(* IEC 61131-3 sources: SRCI_CLIENT_PLC/RobotLibrary/Library/Structures/DatenAndTime, 4 files *)

(* ---- IEC_DATE.st ---- *)
/// Date in the format days since 1990.01.01
TYPE IEC_DATE : UINT;
// -------------------------------------------------------------------------
//  SRCI Robot Library
// -------------------------------------------------------------------------
//
//  Object:      IEC_DATE
//  Author:      Thorsten Brach
//  Date:        2024-06-01
//
//  Description:
//
//
//  Copyright:
//    (C) 2024 Thorsten Brach. All rights reserved
//             Licensed under the MIT License.
//
//  Disclaimer:
//    This project is provided without any guarantee and can be used for
//    private and commercial purposes. Any use is at the user’s
//    own risk and responsibility.
//
// -------------------------------------------------------------------------
END_TYPE

(* ---- IEC_TIME.st ---- *)
/// Time in the clients time zone in the format milliseconds since start of day
TYPE IEC_TIME : TIME_OF_DAY;
// -------------------------------------------------------------------------
//  SRCI Robot Library
// -------------------------------------------------------------------------
//
//  Object:      IEC_TIME
//  Author:      Thorsten Brach
//  Date:        2024-06-01
//
//  Description:
//
//
//  Copyright:
//    (C) 2024 Thorsten Brach. All rights reserved
//             Licensed under the MIT License.
//
//  Disclaimer:
//    This project is provided without any guarantee and can be used for
//    private and commercial purposes. Any use is at the user’s
//    own risk and responsibility.
//
// -------------------------------------------------------------------------
END_TYPE

(* ---- IEC_TIMESTAMP.st ---- *)
TYPE IEC_TIMESTAMP :
// -------------------------------------------------------------------------
//  SRCI Robot Library
// -------------------------------------------------------------------------
//
//  Object:      IEC_TimeStamp
//  Author:      Thorsten Brach
//  Date:        2024-06-11
//
//  Description:
//
//
//  Copyright:
//    (C) 2024 Thorsten Brach. All rights reserved
//             Licensed under the MIT License.
//
//  Disclaimer:
//    This project is provided without any guarantee and can be used for
//    private and commercial purposes. Any use is at the user’s
//    own risk and responsibility.
//
// -------------------------------------------------------------------------
STRUCT
  /// Date
  IEC_DATE : IEC_DATE;
  /// Time
  IEC_TIME : IEC_TIME;
END_STRUCT
END_TYPE

(* ---- SystemTime.st ---- *)
TYPE SystemTime :
// -------------------------------------------------------------------------
//  SRCI Robot Library
// -------------------------------------------------------------------------
//
//  Object:      SystemTime
//  Author:      Thorsten Brach
//  Date:        2025-01-11
//
//  Description:
//
//
//  Copyright:
//    (C) 2025 Thorsten Brach. All rights reserved
//             Licensed under the MIT License.
//
//  Disclaimer:
//    This project is provided without any guarantee and can be used for
//    private and commercial purposes. Any use is at the user’s
//    own risk and responsibility.
//
// -------------------------------------------------------------------------
STRUCT
  /// Date of the system
  SystemDate : DATE;
  /// Time of the system
  SystemTime : TOD;
END_STRUCT
END_TYPE
